(* IEC 61131-3 sources: SemantiST/compiler/intake/normalize/probes/scl-local-prefix, 2 files *)

(* ---- original.st ---- *)
FUNCTION SQUARE : INT
VAR_INPUT
    X : INT;
END_VAR
#SQUARE := #X * #X;
END_FUNCTION

FUNCTION main : DINT
printf('%d$N', SQUARE(3));
main := 0;
END_FUNCTION

(* ---- rewritten.st ---- *)
FUNCTION SQUARE : INT
VAR_INPUT
    X : INT;
END_VAR
SQUARE := X * X;
END_FUNCTION

FUNCTION main : DINT
printf('%d$N', SQUARE(3));
main := 0;
END_FUNCTION
